(* IEC 61131-3 sources: HappyLearnCodesys/content/softmotion/CNC02_online, 3 files *)

(* ---- GVL_Globale_Variablen.st ---- *)
VAR_GLOBAL
	g_x: REAL:=100;
	g_y:REAL:=50;
END_VAR

(* ---- Ipo.st ---- *)
PROGRAM Ipo
VAR
	trafo: SMC_TRAFO_Gantry2;
	p1,p2: SMC_ControlAxisByPos;
	trafof: SMC_TRAFOF_Gantry2;
	smci: SMC_Interpolator;
	mcp1, mcp2: MC_Power;
END_VAR

(* ---- Path.st ---- *)
PROGRAM Path
VAR
	dec: SMC_NCDecoder;
	checkVel: SMC_CheckVelocities;
	buf: ARRAY[0..99] OF SMC_GEOINFO;
END_VAR
